(* IEC 61131-3 sources: volt/packages/volt-lsp-iec/test-corpus/CodesysTestProject/Device/Plc Logic/Application/Library Manager/Analyzation, 8 files *)

(* ---- EXPRESSIONRESULT.dut ---- *)
TYPE EXPRESSIONRESULT :
STRUCT
	NAME : STRING(STRING_LENGTH_EXP);
	ADDRESS : STRING(STRING_LENGTH_ADDRESS);
	COMMENT : STRING(STRING_LENGTH_COMMENT);
	VALUE : BOOL;
	FAILED : BOOL;
END_STRUCT
END_TYPE

(* ---- PARAM.gvl ---- *)
VAR_GLOBAL
	TABLE_UPPER_BOUND : INT := 15;
	STRING_LENGTH_EXP : INT := 255;
	STRING_LENGTH_ADDRESS : INT := 20;
	STRING_LENGTH_COMMENT : INT := 255;
	STRING_LENGTH_OUTSTRING : INT := 255;
	TABLE_SHOW_VALID_ITEMS : BOOL := FALSE;
END_VAR

(* ---- APPENDERRORSTRING.pou ---- *)
FUNCTION APPENDERRORSTRING
VAR_IN_OUT
	STROLD : STRING(STRING_LENGTH_EXP);
	STRNEW : STRING(1);
END_VAR
END_FUNCTION

(* ---- CONCATX.pou ---- *)
FUNCTION CONCATX
VAR_IN_OUT
	STR1 : STRING(STRING_LENGTH_EXP);
	STR2 : STRING(1);
END_VAR
END_FUNCTION

(* ---- LENX.pou ---- *)
FUNCTION LENX : INT
VAR_INPUT
	STR : STRING(STRING_LENGTH_EXP);
END_VAR
END_FUNCTION

(* ---- ANALYZEEXPRESSION.pou ---- *)
FUNCTION_BLOCK ANALYZEEXPRESSION
VAR_INPUT
	INPUTEXP : BOOL;
	DOANALYZE : BOOL;
END_VAR
VAR_OUTPUT
	EXPRESULT : BOOL;
	OUTSTRING : STRING(STRING_LENGTH_OUTSTRING);
END_VAR
END_FUNCTION_BLOCK

METHOD ADDSTRING : BOOL
VAR_IN_OUT
	STRIN : STRING;
END_VAR
END_METHOD

METHOD RESET : BOOL
END_METHOD

(* ---- ANALYZEEXPRESSIONCOMBINED.pou ---- *)
FUNCTION_BLOCK ANALYZEEXPRESSIONCOMBINED
VAR_INPUT
	INPUTEXP : BOOL;
	DOANALYZE : BOOL;
END_VAR
VAR_OUTPUT
	EXPRESULT : BOOL;
	OUTTABLE : ARRAY [0..TABLE_UPPER_BOUND] OF ExpressionResult;
	OUTSTRING : STRING(STRING_LENGTH_OUTSTRING);
END_VAR
VAR
	INDEX : INT;
END_VAR
END_FUNCTION_BLOCK

METHOD ADDENTRY : BOOL
VAR_INPUT
	VALUE : BOOL;
	FAILED : BOOL;
END_VAR
VAR_IN_OUT
	NAME : STRING;
	ADDRESS : STRING;
	COMMENT : STRING;
END_VAR
END_METHOD

METHOD ADDSTRING : BOOL
VAR_IN_OUT
	STRIN : STRING;
END_VAR
END_METHOD

METHOD RESET : BOOL
END_METHOD

(* ---- ANALYZEEXPRESSIONTABLE.pou ---- *)
FUNCTION_BLOCK ANALYZEEXPRESSIONTABLE
VAR_INPUT
	INPUTEXP : BOOL;
	DOANALYZE : BOOL;
END_VAR
VAR_OUTPUT
	EXPRESULT : BOOL;
	OUTTABLE : ARRAY [0..TABLE_UPPER_BOUND] OF ExpressionResult;
END_VAR
VAR
	INDEX : INT;
END_VAR
END_FUNCTION_BLOCK

METHOD ADDENTRY : BOOL
VAR_INPUT
	VALUE : BOOL;
	FAILED : BOOL;
END_VAR
VAR_IN_OUT
	NAME : STRING;
	ADDRESS : STRING;
	COMMENT : STRING;
END_VAR
END_METHOD

METHOD RESET : BOOL
END_METHOD
